{attribute 'linkalways'} 
{attribute 'no_explicit_call' := 'This FB is a CLASS and must be accessed using methods or properties'}
{attribute 'enable_dynamic_creation'}
FUNCTION_BLOCK _Array0to3OfDINT EXTENDS ArrayDatatypeBase_1D
VAR CONSTANT
	lBound : DINT := 0;
	uBound : DINT := 3;
END_VAR
VAR
	localData : ARRAY [lBound..uBound] OF DINT;
	activeData : REFERENCE TO ARRAY [lBound..uBound] OF DINT REF= localData;
	elements : ARRAY [lBound..uBound] OF _DINT(0);
	baseType : _DINT(0);
END_VAR

PROPERTY PUBLIC Address : PVOID
GET
Address := ADR(activeData);
END_GET
END_PROPERTY

PROPERTY PUBLIC BaseDatatype : I_Datatype
GET
BaseDatatype := baseType;
END_GET
END_PROPERTY

METHOD PUBLIC ClearReference
VAR_INPUT
END_VAR
activeData REF= localData;
SetElementReference();
END_METHOD

METHOD PUBLIC Clone : I_Datatype
VAR
    pClone : POINTER TO _Array0to3OfDINT;
END_VAR
pClone := __NEW(_Array0to3OfDINT());
pClone^.Value := Value;
Clone := pClone^;
END_METHOD

METHOD FB_init : BOOL
VAR_INPUT
	bInitRetains : BOOL; // if TRUE, the retain variables are initialized (warm start / cold start)
	bInCopyCode : BOOL;  // if TRUE, the instance afterwards gets moved into the copy code (online change)
END_VAR
SetElementReference();
END_METHOD

METHOD PUBLIC MakeReferenceTo
VAR_INPUT
	ReferenceTarget : REFERENCE TO ARRAY [lBound..uBound] OF DINT;
END_VAR
activeData REF= ReferenceTarget;
SetElementReference();
END_METHOD

METHOD PROTECTED OnSerializeArrayValues
VAR_INPUT
	Serializer : I_Serializer;
END_VAR
VAR
	i : DINT;
END_VAR
FOR i := lBound TO uBound DO
	elements[i].SerializeWith(Serializer);
END_FOR
END_METHOD

METHOD PROTECTED SetElementReference
VAR_INPUT
END_VAR
VAR
	i : DINT;
END_VAR
FOR i := lBound TO uBound DO
	elements[i].MakeReferenceTo(activeData[i]);
END_FOR
END_METHOD

PROPERTY PUBLIC Size : UDINT
GET
Size := SIZEOF(activeData);
END_GET
END_PROPERTY

METHOD PROTECTED TryDeserializeArrayValues : BOOL
VAR_INPUT
	Deserializer : I_Deserializer;
	Feedback : I_DeserializerFeedback;
END_VAR
VAR
	failed : BOOL;
	enumerator : I_DeserializerArrayForwardEnumerator;
	i : DINT;
END_VAR
enumerator := Deserializer.GetArrayEnumerator();
i := lBound;

WHILE enumerator.MoveNext() AND i <= uBound AND NOT failed DO
	
	IF NOT elements[i].TryDeserializeFrom(enumerator.Current, Feedback) THEN
		failed := TRUE;
		EXIT;
	END_IF
	i := i + 1;

END_WHILE
enumerator.Dispose();

TryDeserializeArrayValues := NOT failed;
END_METHOD

METHOD PUBLIC TryGetElementAsDatatypeByIndex : BOOL
VAR_INPUT
	Index : DINT;
	Destination : REFERENCE TO I_Datatype;
END_VAR
IF Index < lbound OR Index > ubound THEN
	RETURN;
END_IF

Destination := elements[Index];
TryGetElementAsDatatypeByIndex := TRUE;
END_METHOD

METHOD PUBLIC TryGetLowerBound : BOOL
VAR_INPUT
	Dimention : UDINT;
	Destination : REFERENCE TO DINT;
END_VAR
IF Dimention = 1 THEN
	Destination := lBound;
	TryGetLowerBound := TRUE;
END_IF
END_METHOD

METHOD PUBLIC TryGetUpperBound : BOOL
VAR_INPUT
	Dimention : UDINT;
	Destination : REFERENCE TO DINT;
END_VAR
IF Dimention = 1 THEN
	Destination := uBound;
	TryGetUpperBound := TRUE;
END_IF
END_METHOD

METHOD TryMakeReferenceTo : BOOL
VAR_INPUT
	Target : I_Datatype;
END_VAR
VAR
	pTargetData : POINTER TO ARRAY [lBound..uBound] OF DINT;
END_VAR
IF NOT IsEquivalentTo(Target) THEN
	RETURN;
END_IF

pTargetData := Target.Address;
activeData REF= pTargetData^;
SetElementReference();
TryMakeReferenceTo := TRUE;
END_METHOD

PROPERTY PUBLIC Value : REFERENCE TO ARRAY [lBound..uBound] OF DINT;
GET
Value ref= activeData;
END_GET
END_PROPERTY

END_FUNCTION_BLOCK

(* stored: Version 1.1.0.1, ProductVersion 3.1.4024.13
   POU _Array0to3OfDINT: Id {64a20a04-94cb-03b2-2a14-f0500ee8ce46}, SpecialFunc None
   Folder Core: Id {8c43b7f1-7fc4-0575-0878-7b1736587bd0}
   Folder Constructor: Id {aa8f9448-f48d-0c34-25ca-f6e68580effb}
   Folder Protected: Id {62143fbf-b4a5-0a08-3acd-76f196378771}
   Folder Customize: Id {7086d3e1-f8ff-01a0-121e-4531e80989d8}
   Property Address: Id {df49b803-c0bd-09c0-135c-6e99b4283be0}
   Get Get: Id {e2c43bca-f08e-0756-2fba-2e7b599bc58d}
   Property BaseDatatype: Id {78ee7d72-dc7b-0189-12b3-ccfea76287cc}
   Get Get: Id {2f1b7f78-c5c3-052e-2a6e-c012c1f6284d}
   Method ClearReference: Id {be1abfab-6b05-0f97-2d8d-b147117b9725}
   Method Clone: Id {3eeb34a1-f8f1-07a3-1aaa-bf7bd3a1726f}
   Method FB_init: Id {13208242-971d-082f-0d50-dda352b4d3b2}
   Method MakeReferenceTo: Id {0883f8ed-e936-019f-02b6-3c5ede4e5518}
   Method OnSerializeArrayValues: Id {7e795148-93d6-082c-3b02-5459f02f0159}
   Method SetElementReference: Id {831e087a-9af2-0a0b-0b6f-96c0b8ae3e14}
   Property Size: Id {d606d92d-8158-0c8a-24d0-976f6d1dc242}
   Get Get: Id {778403c3-e995-0069-181d-86bde3de7c7f}
   Method TryDeserializeArrayValues: Id {99bd456f-2384-0d40-1dbe-28a354944143}
   Method TryGetElementAsDatatypeByIndex: Id {3ab1d446-d473-04da-300c-54f21e140de0}
   Method TryGetLowerBound: Id {05cc96b2-4443-00f7-3c9f-30cfd88c5d57}
   Method TryGetUpperBound: Id {c7356bbc-179f-0bed-28a3-c6240910031f}
   Method TryMakeReferenceTo: Id {64093090-93ca-0771-0ae4-b7f39e4c39d5}
   Property Value: Id {69a4f9fe-17e0-0f0c-3644-8e604e6734fe}
   Get Get: Id {e3e86e7b-b012-08e6-3328-6f4e06c3e183} *)
